Fanuc KAREL source: IO0203.KL

PROGRAM IO0203
%NOLOCKGROUP
ROUTINE RTEST
VAR
L1 : ARRAY[3] OF INTEGER;L2 : XYZWPR
L3 : JOINTPOS9
L4 : POSITION
A:BOOLEAN
S1:INTEGER
B:REAL
C:BOOLEAN
D:REAL
BEGIN
--
--
A=TRUE
L1[1]=2
C=TRUE
D=1.0
SET_JPOS_REG(1,L3,S1,1)
END RTEST
BEGIN
RTEST
END IO0203
